(* IEC 61131-3 sources: PortalRobot/Portal_robot/Device/application/ST/ST_POINT_MANAGER, 8 files *)

(* ---- E_POINT_MANAGER_STATE.st ---- *)
{attribute 'qualified_only'}
{attribute 'strict'}
TYPE E_POINT_MANAGER_STATE :
(
	IDLE,
	SELECT_POINT,
	CHECK_VEL_FACTOR,
	CHECK_ZONE,
	CHECK_ALL
);
END_TYPE

(* ---- ST_POINT_FAULT_REQUEST.st ---- *)
TYPE ST_POINT_FAULT_REQUEST :
STRUCT
	xEnabled        : BOOL; // Глобальное разрешение диагностической инъекции
	xXOutOfLimit    : BOOL; // Импульс проверки точки с недопустимой координатой X
	xYOutOfLimit    : BOOL; // Импульс проверки точки с недопустимой координатой Y
	xZOutOfLimit    : BOOL; // Импульс проверки точки с недопустимой координатой Z
	xInvalidVelocity: BOOL; // Импульс проверки точки с недопустимой скоростью
END_STRUCT
END_TYPE

(* ---- ST_POINT_MANAGER.st ---- *)
TYPE ST_POINT_MANAGER :
STRUCT
	Command : ST_POINT_MANAGER_COMMAND; // Команды менеджера точки
	Status  : ST_POINT_MANAGER_STATUS; // Рабочие статусы менеджера точки
	Diag    : ST_POINT_MANAGER_DIAG; // Состояние автомата и допустимые пределы
	Error   : ST_POINT_MANAGER_ERRORS; // Активные и последние ошибки
END_STRUCT
END_TYPE

(* ---- ST_POINT_MANAGER_COMMAND.st ---- *)
TYPE ST_POINT_MANAGER_COMMAND :
STRUCT
	xExecute : BOOL; // Команда проверки заданной точки
END_STRUCT
END_TYPE

(* ---- ST_POINT_MANAGER_DIAG.st ---- *)
TYPE ST_POINT_MANAGER_DIAG :
STRUCT
	eState       : E_POINT_MANAGER_STATE; // Текущее состояние автомата
	lrX_MinLimit : LREAL; // Минимально допустимая координата X
	lrY_MinLimit : LREAL; // Минимально допустимая координата Y
	lrZ_MinLimit : LREAL; // Минимально допустимая координата Z
	lrX_MaxLimit : LREAL; // Максимально допустимая координата X
	lrY_MaxLimit : LREAL; // Максимально допустимая координата Y
	lrZ_MaxLimit : LREAL; // Максимально допустимая координата Z
	xXLimitValid : BOOL; // Software limits оси X включены и образуют корректный диапазон
	xYLimitValid : BOOL; // Software limits оси Y включены и образуют корректный диапазон
	xZLimitValid : BOOL; // Software limits оси Z включены и образуют корректный диапазон
	stWarning    : ST_WARNING_EVENT; // Последнее предупреждение менеджера точек
END_STRUCT
END_TYPE

(* ---- ST_POINT_MANAGER_ERROR.st ---- *)
TYPE ST_POINT_MANAGER_ERROR :
STRUCT
	X_OUT_OF_LIMIT : BOOL; // Координата X находится вне допустимой зоны
	Y_OUT_OF_LIMIT : BOOL; // Координата Y находится вне допустимой зоны
	Z_OUT_OF_LIMIT : BOOL; // Координата Z находится вне допустимой зоны
	INVALID_VEL    : BOOL; // Коэффициент скорости задан неверно
	X_LIMIT_CONFIG_INVALID : BOOL; // Software limits оси X отключены или заданы некорректно
	Y_LIMIT_CONFIG_INVALID : BOOL; // Software limits оси Y отключены или заданы некорректно
	Z_LIMIT_CONFIG_INVALID : BOOL; // Software limits оси Z отключены или заданы некорректно
	POINT_NOT_CONFIGURED : BOOL; // Инженерная точка ещё не сохранена редактором
END_STRUCT
END_TYPE

(* ---- ST_POINT_MANAGER_ERRORS.st ---- *)
TYPE ST_POINT_MANAGER_ERRORS :
STRUCT
	dwErrorActive : DWORD; // Битовая маска активных ошибок
	dwErrorLast   : DWORD; // Битовая маска последних ошибок
	dwAlarmActive : DWORD; // Собственные аварии менеджера точек для общего журнала
	stErrorActive : ST_POINT_MANAGER_ERROR; // Расшифровка активных ошибок
	stErrorLast   : ST_POINT_MANAGER_ERROR; // Расшифровка последних ошибок
END_STRUCT
END_TYPE

(* ---- ST_POINT_MANAGER_STATUS.st ---- *)
TYPE ST_POINT_MANAGER_STATUS :
STRUCT
	xBusy    : BOOL; // Выполняется проверка точки
	xDone    : BOOL; // Проверка точки завершена
	xInvalid : BOOL; // Точка содержит недопустимые параметры
END_STRUCT
END_TYPE
